// TIA Portal V21 export
FUNCTION_BLOCK "LineSafety"   // FB1, F_FBD
{ S7_Optimized_Access := 'TRUE' }
// Main safety block of the line's F-runtime group.
   VAR
      latched : Bool;
   END_VAR
BEGIN

REGION Network 1: Release
   // Released while start is pressed and the door is closed.
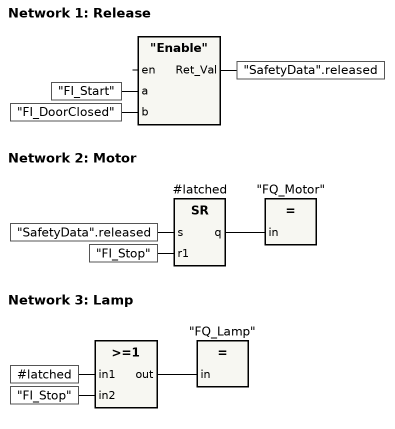
   "SafetyData".released := "Enable"("a" := "FI_Start", "b" := "FI_DoorClosed");
END_REGION

REGION Network 2: Motor
   // Latched on release, dropped by stop.
   IF "SafetyData".released THEN
       #latched := TRUE;   // SR flip-flop
   END_IF;
   IF "FI_Stop" THEN #latched := FALSE; END_IF;
   "FQ_Motor" := #latched;
END_REGION

REGION Network 3: Lamp
   // Lit while the motor runs or stop is pressed.
   "FQ_Lamp" := #latched OR "FI_Stop";
END_REGION
END_FUNCTION_BLOCK
